// TIA Portal V21 export
// export: Created 2026-11-21T13:31:42.105978Z, ExportSetting WithDefaults, DisplayName Totally Integrated Automation Portal, DisplayVersion V21, DisplayName STEP 7 Professional, DisplayVersion V21, DisplayName STEP 7 Safety, DisplayVersion V21, DisplayName Tech WebApplication, DisplayVersion V21, DisplayName WinCC Basic/Comfort/Advanced, DisplayVersion V21, DisplayName WinCC Unified, DisplayVersion V21
VAR_GLOBAL   // PLC tag table "IO"
   Go AT %I0.0 : Bool;   // Carriage start
   Jammed AT %I0.1 : Bool;   // Carriage jammed
   Brake AT %Q0.0 : Bool;   // Carriage brake
   Pointer AT %MD20 : DWord;   // Pointer for indirect access
END_VAR
